(*
SPDX-FileCopyrightText: © 2026 Oleksandr Tiutyk <trofimich@gmail.com>
SPDX-License-Identifier: MIT
License: https://opensource.org/license/mit
*)

(*!
<summary>Checks that a bound TaskStopReason view observes changes to its backing data.</summary>
<description>
Exercises all defined values through the same view in one call. The backing data and view are local to the call.
</description>
*)

{attribute 'no_explicit_call' := 'do not call this function block directly'}
FUNCTION_BLOCK BoundTaskStopReasonTest EXTENDS TOF_Testing.SingleCycleTest
VAR_STAT
	{attribute 'hide'}
	_ClassName : STRING := __POUNAME();
END_VAR

//! <summary>Sets each backing value and checks the corresponding value and flags.</summary>
METHOD PROTECTED ExecuteTest
VAR
	backingValue : TOF_Tasks.TASK_STOP_REASON;
	stopMessage : TOF_Core.ERROR_MESSAGE;
	view : TOF_Tasks.TaskStopReason(stopReason := backingValue, stopReasonMessage := stopMessage);
END_VAR
backingValue := TOF_Tasks.TASK_STOP_REASON.WORK_DONE;
stopMessage := "initial message";
Assert.ThatBool(
	actual := view.Value = TOF_Tasks.TASK_STOP_REASON.WORK_DONE,
	message := "Value must track WORK_DONE"
).IsTrue();
Assert.ThatBool(actual := view.WorkDone, message := "WorkDone must be true for WORK_DONE").IsTrue();
Assert.ThatBool(actual := view.Failure, message := "Failure must be false for WORK_DONE").IsFalse();
Assert.ThatBool(actual := view.ExternalCancel, message := "ExternalCancel must be false for WORK_DONE").IsFalse();
Assert.ThatBool(actual := view.InternalAbort, message := "InternalAbort must be false for WORK_DONE").IsFalse();
Assert.ThatBool(actual := __ISVALIDREF(view.Message), message := "Message must be bound for WORK_DONE").IsTrue();

IF __ISVALIDREF(view.Message) THEN
	Assert.ThatBool(
		actual := view.Message = "initial message",
		message := "Message must match the backing text for WORK_DONE"
	).IsTrue();
END_IF

backingValue := TOF_Tasks.TASK_STOP_REASON.FAILURE;
stopMessage := "diagnostic failure";
Assert.ThatBool(
	actual := view.Value = TOF_Tasks.TASK_STOP_REASON.FAILURE,
	message := "Value must track FAILURE"
).IsTrue();
Assert.ThatBool(actual := view.Failure, message := "Failure must be true for FAILURE").IsTrue();
Assert.ThatBool(actual := view.WorkDone, message := "WorkDone must be false for FAILURE").IsFalse();
Assert.ThatBool(actual := view.ExternalCancel, message := "ExternalCancel must be false for FAILURE").IsFalse();
Assert.ThatBool(actual := view.InternalAbort, message := "InternalAbort must be false for FAILURE").IsFalse();
Assert.ThatBool(actual := __ISVALIDREF(view.Message), message := "Message must be bound for FAILURE").IsTrue();

IF __ISVALIDREF(view.Message) THEN
	Assert.ThatBool(
		actual := view.Message = "diagnostic failure",
		message := "Message must match the backing text for FAILURE"
	).IsTrue();
END_IF

backingValue := TOF_Tasks.TASK_STOP_REASON.EXTERNAL_CANCEL;
Assert.ThatBool(
	actual := view.Value = TOF_Tasks.TASK_STOP_REASON.EXTERNAL_CANCEL,
	message := "Value must track EXTERNAL_CANCEL"
).IsTrue();
Assert.ThatBool(actual := view.ExternalCancel, message := "ExternalCancel must be true for EXTERNAL_CANCEL").IsTrue();
Assert.ThatBool(actual := view.WorkDone, message := "WorkDone must be false for EXTERNAL_CANCEL").IsFalse();
Assert.ThatBool(actual := view.Failure, message := "Failure must be false for EXTERNAL_CANCEL").IsFalse();
Assert.ThatBool(actual := view.InternalAbort, message := "InternalAbort must be false for EXTERNAL_CANCEL").IsFalse();

backingValue := TOF_Tasks.TASK_STOP_REASON.INTERNAL_ABORT;
Assert.ThatBool(
	actual := view.Value = TOF_Tasks.TASK_STOP_REASON.INTERNAL_ABORT,
	message := "Value must track INTERNAL_ABORT"
).IsTrue();
Assert.ThatBool(actual := view.InternalAbort, message := "InternalAbort must be true for INTERNAL_ABORT").IsTrue();
Assert.ThatBool(actual := view.WorkDone, message := "WorkDone must be false for INTERNAL_ABORT").IsFalse();
Assert.ThatBool(actual := view.Failure, message := "Failure must be false for INTERNAL_ABORT").IsFalse();
Assert.ThatBool(actual := view.ExternalCancel, message := "ExternalCancel must be false for INTERNAL_ABORT").IsFalse();
END_METHOD

//! <summary>Borrows the concrete class name. Callers must not modify the returned storage.</summary>
{attribute 'monitoring' := 'call'}
PROPERTY ClassName : REFERENCE TO STRING
GET
ClassName REF= _ClassName;
END_GET
END_PROPERTY

//! <summary>Borrows the compiler-initialized namespace name. Callers must not modify the returned storage.</summary>
{attribute 'monitoring' := 'call'}
PROPERTY NamespaceName : REFERENCE TO STRING
GET
NamespaceName REF= CurrentNamespace.Name;
END_GET
END_PROPERTY

//! <summary>Reports the complete concrete instance size in bytes.</summary>
{attribute 'monitoring' := 'call'}
PROPERTY SelfSize : ULINT
GET
SelfSize := XSIZEOF(THIS^);
END_GET
END_PROPERTY

END_FUNCTION_BLOCK

(* stored: Version 1.1.0.1
   POU BoundTaskStopReasonTest: Id {8e762fbd-f9b4-4f49-84f1-3e6b0340a776}, SpecialFunc None
   Method ExecuteTest: Id {897548ec-ee71-4a70-9d13-c78c1267fc80}
   Property ClassName: Id {8be397be-f8fe-4a75-bc7b-d47761f49846}
   Get Get: Id {f8a9d59c-90ee-4fe7-9d6b-be4446a69845}
   Property NamespaceName: Id {546fe4b3-b7bf-453d-8171-10a2ae552453}
   Get Get: Id {e2c745ee-ebdc-4fec-aa60-2fa910c2fbda}
   Property SelfSize: Id {5fb8c2c9-d014-4f3e-a806-fb10cd9a62a0}
   Get Get: Id {8373f6e7-73c7-452b-9eb6-d756b90d7385} *)
